// Parameters of FB TWOHAND.
TYPE
ST_SafeTwoHandParameters :
STRUCT
    Twohand1MakeContact : BOOL;
    Twohand2MakeContact : BOOL;
    Twohand3MakeContact : BOOL;
    Twohand4MakeContact : BOOL;
    DiscrepancyTime1 : TIME; // Twohand1 / Twohand2
    DiscrepancyTime2 : TIME; // Twohand3 / Twohand4
    HandDiscrepancyTime : TIME; // max time between actuation of the two hands (max 2500 ms). T#0S disables
    SafeInputsAfterDiscError : BOOL; // Safety Editor checkbox 'Safe Inputs after Disc Error', FALSE for a new block:
        // TRUE makes both channels of the pair that raised a discrepancy error return to the safe state together
        // before ErrAck can clear it
END_STRUCT
END_TYPE

(* stored: Version 1.1.0.1
   DUT ST_SafeTwoHandParameters: Id {b88544d9-b726-539b-a312-7f8941f8befd} *)
